Fanuc KAREL source: KT00458.KL

PROGRAM KT00458
%NOLOCKGROUP
VAR
  P1: POSITION
  P2: JOINTPOS
  OUT: BOOLEAN
BEGIN
  OUT = P1 >= P2
END KT00458
